// TIA Portal V20 export
Screen "190FX1Layout"  1276x673
  ScreenItem "Line_Header_X0_Y64" at 0,64 size 1276x0  Type=HmiLine
  ScreenItem "permanentareaborderrectangle" at 0,0 size 0x0  Type=HmiRectangle
  ScreenItem "Button_Back" at 2,2 size 90x60  Type=HmiButton
  ScreenItem "Move_Legend" at 1182,2 size 90x60  Type=HmiButton
  ScreenItem "Fusszeile_Button_ManualOPMode1_2" at 279,2 size 90x60  Type=HmiButton
  ScreenItem "文本域_3" at 1107,71 size 139x22  Type=HmiTextBox
  ScreenItem "文本域_1" at 1107,160 size 156x23  Type=HmiTextBox
  ScreenItem "文本域_2" at 1107,246 size 135x23  Type=HmiTextBox
  ScreenItem "文本域_22" at 1125,476 size 104x23  Type=HmiTextBox
  ScreenItem "面板容器_2" at 1090,4 size 88x58  Type=HmiFaceplateContainer
  ScreenItem "OPMode1_Blocked" at 1164,6 size 14x14  Type=HmiGraphicView
  ScreenItem "OPMode4_Foreground_Blocked" at 1089,2 size 88x58  Type=HmiGraphicView
  ScreenItem "Fusszeile_Button_ManualOPMode1_1" at 95,2 size 90x60  Type=HmiButton
  ScreenItem "文本域_4" at 1107,330 size 139x22  Type=HmiTextBox
  ScreenItem "Button_Back_1" at 1180,606 size 90x60  Type=HmiButton
  ScreenItem "Fusszeile_Button_ManualOPMode1_3" at 187,2 size 90x60  Type=HmiButton
  ScreenItem "Fusszeile_Button_ManualOPMode1_4" at 997,2 size 90x60  Type=HmiButton
  ScreenItem "Fusszeile_Button_ManualOPMode1_5" at 902,1 size 90x60  Type=HmiButton
  ScreenItem "文本域_14" at 936,-172 size 140x40  Type=HmiTextBox
  ScreenItem "Title_ScreenOverview_X390_Y2_1" at 384,5 size 510x57  Type=HmiTextBox
  ScreenItem "Faceplate container_1" at 229,510 size 61x45  Type=HmiFaceplateContainer
  ScreenItem "Faceplate container_4" at 27,219 size 59x43  Type=HmiFaceplateContainer
  ScreenItem "Graphic view_1" at 19,230 size 860x259  Type=HmiGraphicView
  ScreenItem "Line_9" at 558,162 size 94x182  Type=HmiLine
  ScreenItem "Line_2" at 702,237 size 20x91  Type=HmiLine
  ScreenItem "Line_5" at 752,169 size 73x168  Type=HmiLine
  ScreenItem "Line_17" at 90,242 size 189x81  Type=HmiLine
  ScreenItem "Line_6" at 751,326 size 173x47  Type=HmiLine
  ScreenItem "Line_10" at 632,412 size 84x81  Type=HmiLine
  ScreenItem "Line_13" at 729,414 size 25x80  Type=HmiLine
  ScreenItem "Line_1" at 536,375 size 127x111  Type=HmiLine
  ScreenItem "Line_18" at 262,417 size 17x71  Type=HmiLine
  ScreenItem "Line_16" at 122,341 size 33x138  Type=HmiLine
  ScreenItem "面板容器_4" at 596,518 size 56x46  Type=HmiFaceplateContainer
  ScreenItem "文本域_6" at 45,477 size 140x40  Type=HmiTextBox
  ScreenItem "文本域_7" at 206,487 size 100x20  Type=HmiTextBox
  ScreenItem "文本域_8" at 454,487 size 100x40  Type=HmiTextBox
  ScreenItem "文本域_9" at 574,495 size 100x20  Type=HmiTextBox
  ScreenItem "文本域_10" at 700,494 size 140x40  Type=HmiTextBox
  ScreenItem "文本域_12" at 918,300 size 100x40  Type=HmiTextBox
  ScreenItem "文本域_13" at 502,98 size 140x20  Type=HmiTextBox
  ScreenItem "文本域_15" at 918,412 size 140x40  Type=HmiTextBox
  ScreenItem "文本域_17" at 7,196 size 100x20  Type=HmiTextBox
  ScreenItem "文本域_18" at 652,176 size 100x20  Type=HmiTextBox
  ScreenItem "文本域_20" at 766,98 size 140x20  Type=HmiTextBox
  ScreenItem "Line_11" at 378,190 size 45x115  Type=HmiLine
  ScreenItem "Line_4" at 235,187 size 179x140  Type=HmiLine
  ScreenItem "Line_12" at 777,236 size 144x103  Type=HmiLine
  ScreenItem "Line_19" at 777,402 size 136x24  Type=HmiLine
  ScreenItem "文本域_26" at 918,176 size 140x40  Type=HmiTextBox
  ScreenItem "文本域_11" at 908,515 size 140x20  Type=HmiTextBox
  ScreenItem "Line_3" at 757,411 size 148x112  Type=HmiLine
  ScreenItem "Faceplate container_2" at 344,510 size 69x45  Type=HmiFaceplateContainer
  ScreenItem "文本域_16" at 329,487 size 100x20  Type=HmiTextBox
  ScreenItem "Line_7" at 408,411 size 156x74  Type=HmiLine
  ScreenItem "文本域_19" at 433,179 size 100x20  Type=HmiTextBox
  ScreenItem "Line_8" at 488,246 size 81x78  Type=HmiLine
  ScreenItem "文本域_23" at 281,98 size 140x40  Type=HmiTextBox
  ScreenItem "文本域_21" at 128,98 size 140x40  Type=HmiTextBox
  ScreenItem "面板容器_8" at 130,139 size 144x51  Type=HmiFaceplateContainer
  ScreenItem "面板容器_11" at 282,137 size 150x51  Type=HmiFaceplateContainer
  ScreenItem "面板容器_5" at 45,518 size 143x50  Type=HmiFaceplateContainer
  ScreenItem "面板容器_10" at 512,120 size 153x58  Type=HmiFaceplateContainer
  ScreenItem "面板容器_9" at 908,534 size 148x58  Type=HmiFaceplateContainer
  ScreenItem "面板容器_15" at 921,216 size 149x54  Type=HmiFaceplateContainer
  ScreenItem "面板容器_6" at 921,454 size 149x54  Type=HmiFaceplateContainer
  ScreenItem "Faceplate container_6" at 938,340 size 59x45  Type=HmiFaceplateContainer
  ScreenItem "面板容器_20" at 700,537 size 150x51  Type=HmiFaceplateContainer
  ScreenItem "Faceplate container_7" at 474,529 size 59x45  Type=HmiFaceplateContainer
  ScreenItem "文本域_5" at -1,82 size 120x40  Type=HmiTextBox
  ScreenItem "文本域_27" at -1,126 size 120x40  Type=HmiTextBox
  ScreenItem "LSicar_Valve8Pos_LeftHomeRightWork_WithPB_5" at 1099,95 size 160x53  Type=HmiFaceplateContainer
  ScreenItem "LSicar_Valve8Pos_LeftHomeRightWork_WithPB_1" at 1099,183 size 160x53  Type=HmiFaceplateContainer
  ScreenItem "面板容器_22" at 1062,509 size 96x32  Type=HmiFaceplateContainer
  ScreenItem "面板容器_23" at 1172,509 size 96x32  Type=HmiFaceplateContainer
  ScreenItem "LSicar_Valve8Pos_LeftHomeRightWork_WithPB_2" at 1099,271 size 160x53  Type=HmiFaceplateContainer
  ScreenItem "LSicar_Valve8Pos_LeftHomeRightWork_WithPB_3" at 1099,359 size 160x53  Type=HmiFaceplateContainer
  ScreenItem "面板容器_7" at 766,120 size 148x58  Type=HmiFaceplateContainer
  ScreenItem "Faceplate container_5" at 453,202 size 59x43  Type=HmiFaceplateContainer
  ScreenItem "Faceplate container_3" at 670,197 size 59x45  Type=HmiFaceplateContainer
  ScreenItem "Button_Back_2" at 8,606 size 90x60  Type=HmiButton
  ScreenItem "Button_Back_3" at 122,606 size 90x60  Type=HmiButton
